Staubli VAL3: appStart.pjx

--- appStart.pjx ---
Parameters version=s8.15.3Cs9_BS3337 stackSize=200000 millimeterUnit=true
Program file=start.pgx
Program file=stop.pgx
Program file=Page_AppStart.pgx
Program file=taskHmi.pgx
Program file=_clickProfile.pgx
Program file=_clickFuncReset.pgx
Data file=appStart.dtx

--- appStart.dtx ---
public string sAppName = "MainApp"
public string sDbId = ""
public string sRobotModel
public string sRobotSN
public string sCtrlSN
public string sProfile
public string sProfileRaw
public string sLogin[2]
  [0] = "operator"
  [1] = "programmer"
public string sRoleName[2]
  [0] = "生产员"
  [1] = "工程师"
public bool bFunc[9]
public string sFuncBg[9]
  [0] = "#DCDCDC"
  [1] = "#DCDCDC"
  [2] = "#DCDCDC"
  [3] = "#DCDCDC"
  [4] = "#DCDCDC"
  [5] = "#DCDCDC"
  [6] = "#DCDCDC"
  [7] = "#DCDCDC"
  [8] = "#DCDCDC"
public bool bBtnPressed[9]

--- start.pgx ---
program start()
begin
  //应用入口。SRS 下载后在“应用管理”里设为启动应用即可自动执行。
  //1) 初始化主界面：取设备信息 + 打开页面 + 绑定 9 个功能按钮
  call Page_AppStart()

  //2) 常驻 HMI 任务：刷新角色、同步按钮背景色（优先级低于工艺任务）
  taskCreate "taskHmi",50,taskHmi()

  //3) 主程序作为心跳，不退出
  do
    delay(1)
  until false
end

--- _clickFuncReset.pgx ---
public program _clickFuncReset()
  local num l_nI
begin
  //“全部复位”按钮回调（无参数，供 AppStart.bindings.json 的 callbacks 调用）
  //9 个功能按钮选中态清零，背景色回默认灰
  for l_nI=0 to 8
    bFunc[l_nI]=false
    sFuncBg[l_nI]="#DCDCDC"
  endFor
end

--- _clickProfile.pgx ---
public program _clickProfile()
  local num l_nCur
  local num l_nTarget
  local num l_nRet
  local string l_sPwd
  local string l_sMsg
begin
  //权限图标点击回调（无参数，供 AppStart.bindings.json 的 callbacks 调用）
  //两级角色：0=生产员(operator) 1=工程师(programmer)
  //手册依据：userPageConfirm/userPagePrompt 第81-82页、getProfile/setProfile 第83页

  //1) 判断当前角色
  l_nCur=-1
  if sProfileRaw==sLogin[0]
    l_nCur=0
  elseIf sProfileRaw==sLogin[1]
    l_nCur=1
  endIf

  //2) 目标是"另一个角色"（当前是 staubli/未知时默认切到生产员）
  if l_nCur==0
    l_nTarget=1
  else
    l_nTarget=0
  endIf

  //3) 确认 + 输密码
  l_sMsg="当前："+sProfile+"，是否切换到 "+sRoleName[l_nTarget]+"？"
  if userPageConfirm(l_sMsg)==false
    return
  endIf

  l_sPwd=""
  if userPagePrompt("请输入"+sRoleName[l_nTarget]+"的密码",l_sPwd)==false
    return
  endIf

  //4) 切换并刷新显示名
  l_nRet=setProfile(sLogin[l_nTarget],l_sPwd)
  if l_nRet==0
    sProfileRaw=getProfile()
    sProfile=sProfileRaw
    if sProfileRaw==sLogin[0]
      sProfile=sRoleName[0]
    elseIf sProfileRaw==sLogin[1]
      sProfile=sRoleName[1]
    endIf
  elseIf l_nRet==-1
    userPageAlert("切换失败(-1)：用户未定义，请核对 appStart.dtx 里 sLogin 的登录名")
  elseIf l_nRet==-2
    userPageAlert("切换失败(-2)：密码错误")
  elseIf l_nRet==-3
    userPageAlert("切换失败(-3)：不允许使用 staubli 用户")
  elseIf l_nRet==-4
    userPageAlert("切换失败(-4)：当前是 staubli 用户，不能切换")
  else
    userPageAlert("切换失败，错误码："+toString("",l_nRet))
  endIf
end

--- Page_AppStart.pgx ---
public program Page_AppStart()
  local num l_nRet
begin
  //主界面初始化（只跑一次）：取设备信息 -> 打开页面 -> 绑 9 个功能按钮
  //手册依据：getVersion 第124页、userPage 第75页、userPageBindClick 第78页

  //1) 设备信息
  sRobotModel=getVersion("Arm Type")
  sRobotSN=getVersion("Arm S/N")
  sCtrlSN=getVersion("Controller S/N")

  //2) 权限转两级角色显示名（生产员 / 工程师），原始值另存 sProfileRaw
  //注意：sLogin 里的 "operator"/"programmer" 必须与控制器“用户管理”里实际定义的
  //      profile 名一致，否则 setProfile 返回 -1；现场不同就改 appStart.dtx
  sProfileRaw=getProfile()
  sProfile=sProfileRaw
  if sProfileRaw==sLogin[0]
    sProfile=sRoleName[0]
  elseIf sProfileRaw==sLogin[1]
    sProfile=sRoleName[1]
  endIf

  //3) 打开页面（页面文件是 interface/AppStart.html，名字不带扩展名）
  l_nRet=userPage("AppStart")
  if l_nRet!=0
    userPageAlert("主界面加载失败，请检查 interface/AppStart.html 是否存在")
  endIf

  //4) 9 个功能按钮：点击把对应 bFunc 置 true（不是取反），背景色由 sFuncBg 绑定
  userPageBindClick("AppStart","btn_func1",bFunc[0],true)
  userPageBindClick("AppStart","btn_func2",bFunc[1],true)
  userPageBindClick("AppStart","btn_func3",bFunc[2],true)
  userPageBindClick("AppStart","btn_func4",bFunc[3],true)
  userPageBindClick("AppStart","btn_func5",bFunc[4],true)
  userPageBindClick("AppStart","btn_func6",bFunc[5],true)
  userPageBindClick("AppStart","btn_func7",bFunc[6],true)
  userPageBindClick("AppStart","btn_func8",bFunc[7],true)
  userPageBindClick("AppStart","btn_func9",bFunc[8],true)

  //label（lbl_appname / lbl_model / lbl_sn / lbl_dbid / lbl_profile）的绑定在
  //interface/AppStart.bindings.json 里，这里不要重复绑，否则两处会打架
end

--- stop.pgx ---
program stop()
  local num l_nI
begin
  //应用停止时调用：清掉 9 个功能按钮的选中态，避免下次启动带着上次的状态
  for l_nI=0 to 8
    bFunc[l_nI]=false
    sFuncBg[l_nI]="#DCDCDC"
  endFor
end

--- taskHmi.pgx ---
public program taskHmi()
  local num l_nI
  local bool l_bPrev[9]
begin
  //常驻 HMI 任务：1 秒刷新角色，bFunc 变化时同步按钮背景色
  //注意：循环里必须有 delay()，否则会把控制器 CPU 跑满

  //上电先对齐一次：记录当前选中态并刷新背景色
  for l_nI=0 to 8
    l_bPrev[l_nI]=bFunc[l_nI]
    if bFunc[l_nI]
      sFuncBg[l_nI]="#4CAF50"
    else
      sFuncBg[l_nI]="#DCDCDC"
    endIf
  endFor

  do
    //1) 刷新角色（可能被示教器/MCP 侧改掉），原始值进 sProfileRaw，显示名进 sProfile
    sProfileRaw=getProfile()
    sProfile=sProfileRaw
    if sProfileRaw==sLogin[0]
      sProfile=sRoleName[0]
    elseIf sProfileRaw==sLogin[1]
      sProfile=sRoleName[1]
    endIf

    //2) bFunc 变化时同步背景色：选中 #4CAF50，复位 #DCDCDC
    for l_nI=0 to 8
      if bFunc[l_nI]!=l_bPrev[l_nI]
        l_bPrev[l_nI]=bFunc[l_nI]
        if bFunc[l_nI]
          sFuncBg[l_nI]="#4CAF50"
        else
          sFuncBg[l_nI]="#DCDCDC"
        endIf
      endIf
    endFor

    //3) 让出 CPU，周期 1 秒
    delay(1)
  until false
end
